(*
SPDX-FileCopyrightText: c 2026 Oleksandr Tiutyk <trofimich@gmail.com>
SPDX-License-Identifier: MIT
License: https://opensource.org/license/mit
*)

(*!
<summary>Checks predicate matching, skip, reverse traversal and absence.</summary>
<description>
Borrows a group-owned list reserved for this case. Use from one task at a stable address.
Teardown clears the list before publication.
</description>
*)

{attribute 'no_assign'}
{attribute 'no_explicit_call' := 'do not call this function block directly'}
FUNCTION_BLOCK ListFindTest EXTENDS TOF_Testing.SingleCycleTest
VAR_STAT
	{attribute 'hide'}
	_ClassName : STRING := __POUNAME();
END_VAR
VAR
	_List : TOF_Collections.IList;
	_Predicate : ListStringPredicate;
END_VAR

(*!
<summary>Clears the fixture before the runner publishes the result.</summary>
<description>
Also runs after an unexpected exception interrupts the case.
</description>
*)
METHOD PROTECTED AfterTest
_List.Clear();
END_METHOD

//! <summary>Borrows the concrete class name. Callers must not modify it.</summary>
{attribute 'monitoring' := 'call'}
PROPERTY ClassName : REFERENCE TO STRING
GET
ClassName REF= _ClassName;
END_GET
END_PROPERTY

(*!
<summary>Checks predicate matching, skip, reverse traversal and absence.</summary>
*)
METHOD PROTECTED ExecuteTest
VAR
	values : ARRAY [0..5] OF STRING := ['String0', 'String1', 'String2', 'String3', 'String4', 'String5'];
	found : BOOL;
	index : TOF_Core.DINT_INDEX;
	entry : TOF_Core.GENERIC_VALUE;
END_VAR
_List.AppendCopy(value := values[0]);
_List.AppendCopy(value := values[1]);
_List.AppendCopy(value := values[2]);
_List.AppendCopy(value := values[3]);
_List.AppendCopy(value := values[4]);
_List.AppendCopy(value := values[5]);
_List.AppendCopy(value := values[2]);
_List.AppendCopy(value := values[3]);

_Predicate.Expected := 'String2';

found := _List.FindSingle(predicate := _Predicate, skip := 0, index => index, value => entry);

Assert.ThatBool(
	actual := found AND_THEN index = 2 AND_THEN entry.AsString255() = 'String2',
	message := "Find must return the first match and its value"
).IsTrue();

found := _List.FindSingle(predicate := _Predicate, skip := 1, index => index);

Assert.ThatBool(
	actual := found AND_THEN index = 6,
	message := "Skipping one match must return the second match"
).IsTrue();

found := _List.FindSingle(
	predicate := _Predicate,
	searchDirection := TOF_Core.SEARCH_DIRECTION.FROM_END,
	index => index
);

Assert.ThatBool(
	actual := found AND_THEN index = 6,
	message := "Reverse traversal must find the last occurrence first"
).IsTrue();

found := _List.FindSingle(predicate := _Predicate, skip := 2);

Assert.ThatBool(
	actual := found,
	message := "Skipping both matches must report absence"
).IsFalse();

Assert.ThatDInt(
	actual := _List.Length,
	message := "Find must preserve the list length"
).ToBe(expected := DINT#8);
END_METHOD

(*!
<summary>Binds the list fixture for this case.</summary>
<description>
Stores a borrowed interface without invoking the fixture. The owning group keeps it alive and
reserves it for this case. TestElement initializes the name and parent.
</description>
<param name="name">Display name of this case.</param>
<param name="parent">Group that owns this case.</param>
<param name="list">Required live list reserved for this case.</param>
*)
METHOD FB_init : BOOL
VAR_INPUT
	bInitRetains: BOOL; // TRUE: the retain variables are initialized (reset warm / reset cold)
	bInCopyCode: BOOL; // TRUE: the instance will be copied to the copy code afterward (online change)
	name : WSTRING;
	parent : TOF_Testing.ITestElement;
	list : TOF_Collections.IList;
END_VAR
_List := list;
FB_init := TRUE;
END_METHOD

//! <summary>Borrows the compiler-initialized namespace name. Callers must not modify it.</summary>
{attribute 'monitoring' := 'call'}
PROPERTY NamespaceName : REFERENCE TO STRING
GET
NamespaceName REF= CurrentNamespace.Name;
END_GET
END_PROPERTY

//! <summary>Reports the concrete instance size in bytes.</summary>
{attribute 'monitoring' := 'call'}
PROPERTY SelfSize : ULINT
GET
SelfSize := XSIZEOF(THIS^);
END_GET
END_PROPERTY

END_FUNCTION_BLOCK

(* stored: Version 1.1.0.1, ProductVersion 3.1.4026.21
   POU ListFindTest: Id {21976fa8-b530-46e1-bf48-990a34f9b32d}, SpecialFunc None
   Method AfterTest: Id {4208eb5d-a57a-4362-b11a-842efc9eb921}
   Property ClassName: Id {547bfcb1-5219-4707-8bc5-96d1115e9543}
   Get Get: Id {ff431ede-7d12-44bd-8b3b-8c64a7c9acbf}
   Method ExecuteTest: Id {6eaf83e3-fb36-4b41-bdc6-cb0924cb85d6}
   Method FB_init: Id {9ed88c82-df5e-4979-b07e-ea28c8f693dc}
   Property NamespaceName: Id {bb388751-6825-4574-9d76-95e96d1cc452}
   Get Get: Id {5c759424-53ed-4b30-8416-6e85b4ac3dde}
   Property SelfSize: Id {c1e63185-e73e-459c-8b07-53c69fd7d671}
   Get Get: Id {d6c6f016-2517-47e5-9ced-b7e696671f4b} *)
